Fanuc KAREL source: KT00723.KL

PROGRAM KT00723
%NOLOCKGROUP
VAR
  P1: XYZWPREXT
  P2: XYZWPREXT
  OUT: INTEGER
BEGIN
  P1.X = 1.0
  P2.Y = 2.0
  P1.X = 1.0
  P2.Y = 2.0
  OUT = ARRAY_LEN(P1)
END KT00723
